RoboDK station: hand_motion - lara.rdk

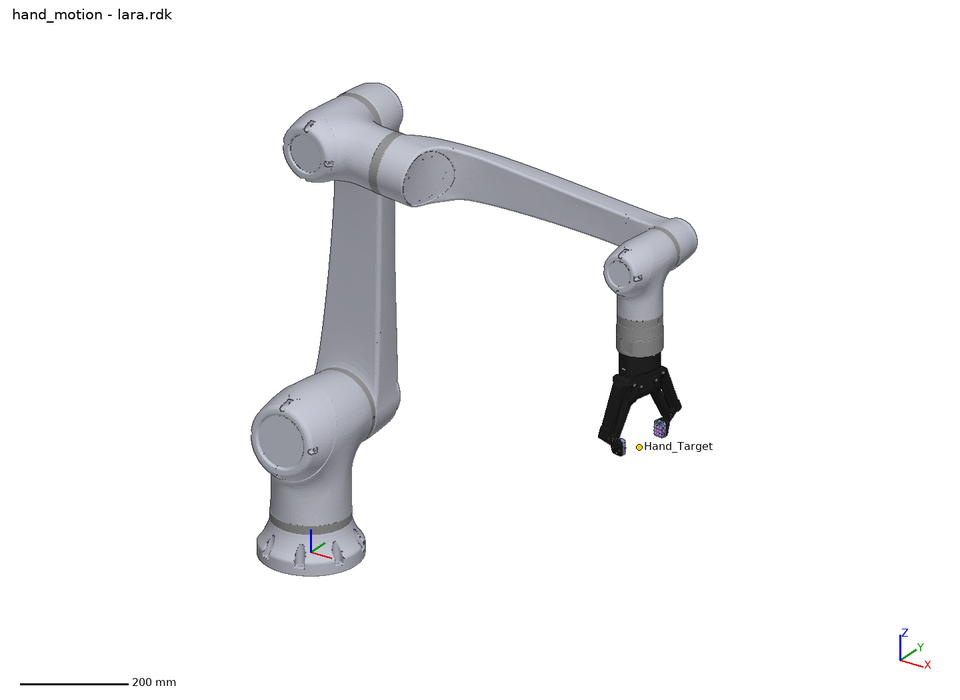
[picture v0: the station drawn from its stored meshes, robots at their saved joint values, targets as dots, program paths as lines]
Station hand_motion (saved by RoboDK 6.0.3). Poses are relative to the parent item; angles as X-Y-Z fixed-axis rotations.
  - frame Neura LARA 8 Base at (0, 0, 0) mm
    - robot Neura LARA 8: 6 axes
        modified DH rows (alpha deg, a mm, theta deg, d mm): 0, 0, 0, 260; -90, 0, -90, 0; 0, 600, -90, 0; -90, 0, 0, 700; 90, 0, 0, 0; -90, 0, 180, 179.5
        joint limits [-180, -135, -155, -180, -180, -360] to [180, 135, 155, 180, 180, 360]; home [0, 0, 90, 0, 90, 0]; saved at [0, 4.031, 90.642, 0, 85.327, 0]
      - tool GAL2_B1.1_CustomerFacing_88mm, TCP at (0, 0, 200) mm, size 75.9 x 197.2 x 204.3 mm, geometry from GAL2_B1.1_CustomerFacing_88mm.STEP
    - target Hand_Target (Cartesian target) at (739.85, 0, 421.99) mm, rotated rx 180 ry 0 rz -180 deg; joints [0, 27.366, 81.033, 0, 71.601, 0] of Neura LARA 8
